// TIA Portal V20 export
// export: Created 2026-10-19T18:41:39.9754622Z, ExportSetting WithDefaults, DisplayName Totally Integrated Automation Portal, DisplayVersion V20 Update 6, DisplayName TIA Portal Openness, DisplayVersion V20 Update 6, DisplayName TIA Portal Version Control Interface, DisplayVersion V20 Update 6, DisplayName SINAMICS Startdrive Advanced, DisplayVersion V20 SP1, DisplayName SINAMICS Startdrive G130, G150, S120, S150, SINAMICS MV, G220, S200, S210, DisplayVersion V20 SP1, DisplayName SINAMICS Startdrive G110M, G120, G120C, G120D, G120P, G115D, DisplayVersion V20 SP1, DisplayName STEP 7 Professional, DisplayVersion V20 Update 6, DisplayName STEP 7 Safety, DisplayVersion V20 Update 2, DisplayName WinCC Basic/Comfort/Advanced, DisplayVersion V20 Update 6, DisplayName WinCC Unified, DisplayVersion V20 Update 6
FUNCTION "FC_CLOCK" : DTL   // FC55, LAD
{ S7_Optimized_Access := 'TRUE' }
VERSION : 0.1
// stored: AutoNumber true, IsIECCheckEnabled false, SetENOAutomatically false, UDAEnableTagReadback false
   VAR_OUTPUT
      CurrentTime : String;
   END_VAR
   VAR_TEMP
      CurrentDTL : DTL;
      RetVal : Int;
      TempString : String;
      strYear : String;
      strMonth : String;
      strDay : String;
      strHour : String;
      strMinute : String;
      strSeconds : String;
   END_VAR
   VAR_TEMP   // added for the SCL form of the ladder/FBD networks
      _w1 : Bool;
      _w2 : Bool;
      _w3 : Bool;
      _w4 : Bool;
      _w5 : Bool;
   END_VAR
BEGIN

REGION Network 1: Read Current Local Time
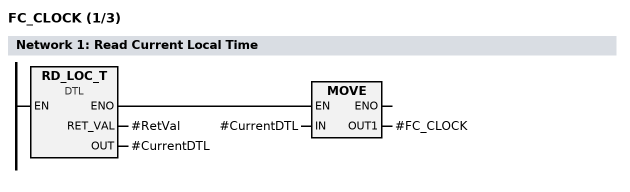
   RUNG wire#powerrail
      { S7_Templates := "date_type := DTL" } RD_LOC_T(RET_VAL => #RetVal, OUT => #CurrentDTL)
      Move(in := #CurrentDTL, out1 => #FC_CLOCK)
   END_RUNG
   // the same network as SCL:
   #RetVal := RD_LOC_T(OUT => #CurrentDTL, ENO => #_w1);
   IF #_w1 THEN #FC_CLOCK := #CurrentDTL; END_IF;
END_REGION

REGION Network 2: Converstion all data to string
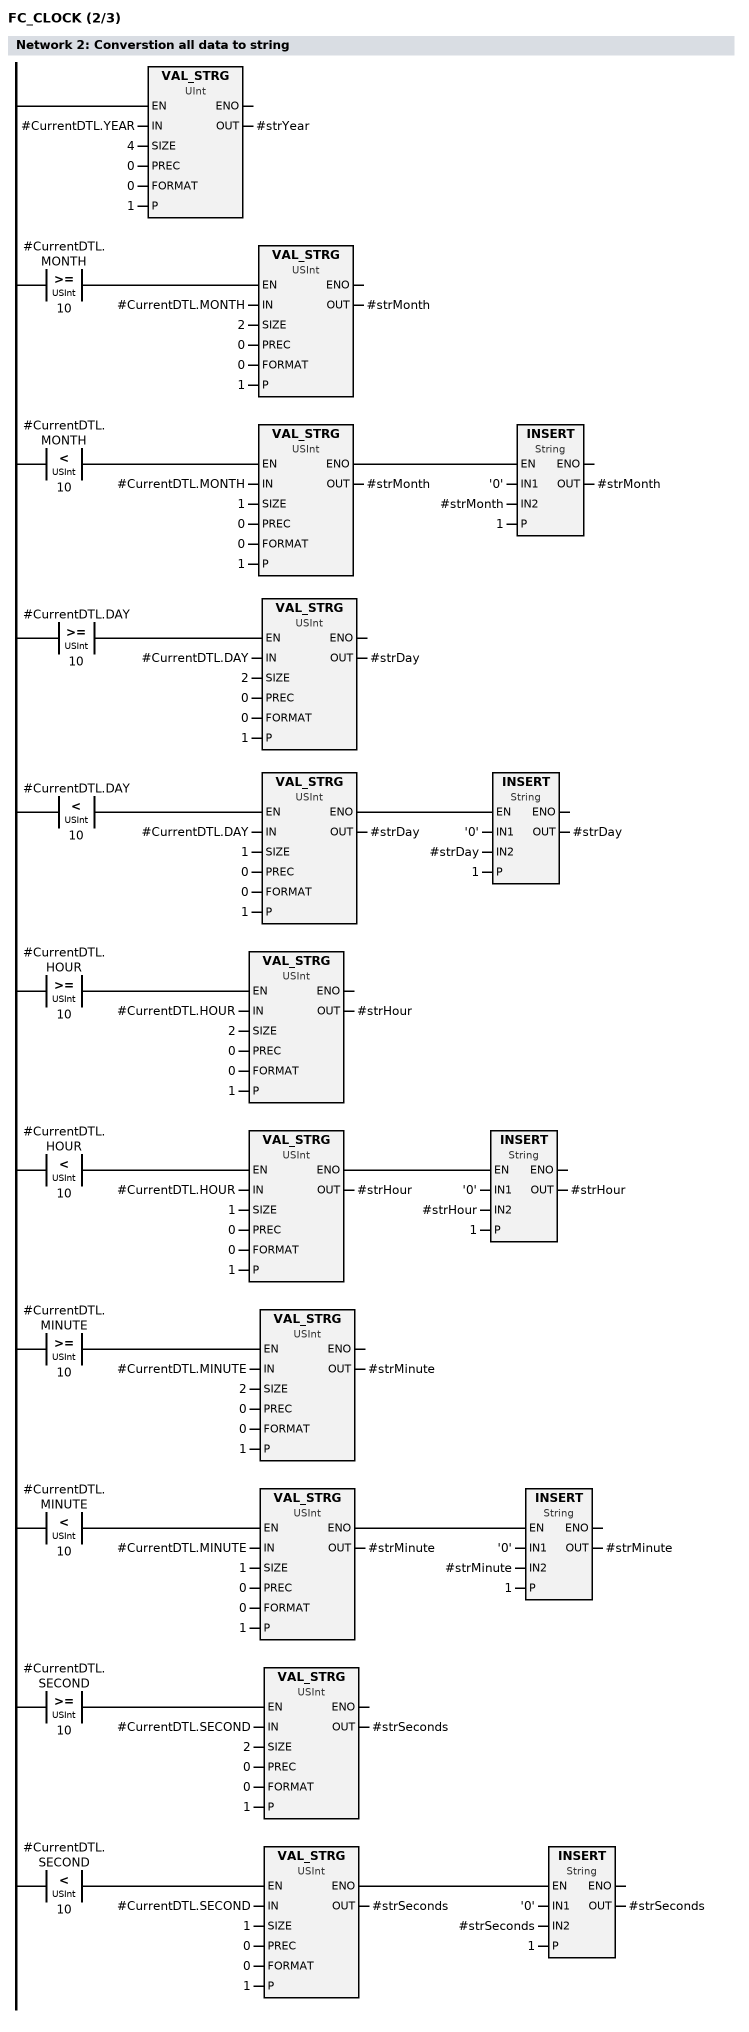
   RUNG wire#powerrail
      { S7_Templates := "[value_type := UInt, str_type := String]" } VAL_STRG(IN := #CurrentDTL.YEAR, SIZE := 4, PREC := 0, FORMAT := 0, P := 1, OUT => #strYear)
   END_RUNG
   RUNG wire#powerrail
      { S7_Templates := "SrcType := USInt" } GE_Contact(in1 := #CurrentDTL.MONTH, in2 := 10)
      { S7_Templates := "[value_type := USInt, str_type := String]" } VAL_STRG(IN := #CurrentDTL.MONTH, SIZE := 2, PREC := 0, FORMAT := 0, P := 1, OUT => #strMonth)
   END_RUNG
   RUNG wire#powerrail
      { S7_Templates := "SrcType := USInt" } LT_Contact(in1 := #CurrentDTL.MONTH, in2 := 10)
      { S7_Templates := "[value_type := USInt, str_type := String]" } VAL_STRG(IN := #CurrentDTL.MONTH, SIZE := 1, PREC := 0, FORMAT := 0, P := 1, OUT => #strMonth)
      { S7_Templates := "str_type := String" } INSERT(IN1 := '0', IN2 := #strMonth, P := 1, OUT => #strMonth)
   END_RUNG
   RUNG wire#powerrail
      { S7_Templates := "SrcType := USInt" } GE_Contact(in1 := #CurrentDTL.DAY, in2 := 10)
      { S7_Templates := "[value_type := USInt, str_type := String]" } VAL_STRG(IN := #CurrentDTL.DAY, SIZE := 2, PREC := 0, FORMAT := 0, P := 1, OUT => #strDay)
   END_RUNG
   RUNG wire#powerrail
      { S7_Templates := "SrcType := USInt" } LT_Contact(in1 := #CurrentDTL.DAY, in2 := 10)
      { S7_Templates := "[value_type := USInt, str_type := String]" } VAL_STRG(IN := #CurrentDTL.DAY, SIZE := 1, PREC := 0, FORMAT := 0, P := 1, OUT => #strDay)
      { S7_Templates := "str_type := String" } INSERT(IN1 := '0', IN2 := #strDay, P := 1, OUT => #strDay)
   END_RUNG
   RUNG wire#powerrail
      { S7_Templates := "SrcType := USInt" } GE_Contact(in1 := #CurrentDTL.HOUR, in2 := 10)
      { S7_Templates := "[value_type := USInt, str_type := String]" } VAL_STRG(IN := #CurrentDTL.HOUR, SIZE := 2, PREC := 0, FORMAT := 0, P := 1, OUT => #strHour)
   END_RUNG
   RUNG wire#powerrail
      { S7_Templates := "SrcType := USInt" } LT_Contact(in1 := #CurrentDTL.HOUR, in2 := 10)
      { S7_Templates := "[value_type := USInt, str_type := String]" } VAL_STRG(IN := #CurrentDTL.HOUR, SIZE := 1, PREC := 0, FORMAT := 0, P := 1, OUT => #strHour)
      { S7_Templates := "str_type := String" } INSERT(IN1 := '0', IN2 := #strHour, P := 1, OUT => #strHour)
   END_RUNG
   RUNG wire#powerrail
      { S7_Templates := "SrcType := USInt" } GE_Contact(in1 := #CurrentDTL.MINUTE, in2 := 10)
      { S7_Templates := "[value_type := USInt, str_type := String]" } VAL_STRG(IN := #CurrentDTL.MINUTE, SIZE := 2, PREC := 0, FORMAT := 0, P := 1, OUT => #strMinute)
   END_RUNG
   RUNG wire#powerrail
      { S7_Templates := "SrcType := USInt" } LT_Contact(in1 := #CurrentDTL.MINUTE, in2 := 10)
      { S7_Templates := "[value_type := USInt, str_type := String]" } VAL_STRG(IN := #CurrentDTL.MINUTE, SIZE := 1, PREC := 0, FORMAT := 0, P := 1, OUT => #strMinute)
      { S7_Templates := "str_type := String" } INSERT(IN1 := '0', IN2 := #strMinute, P := 1, OUT => #strMinute)
   END_RUNG
   RUNG wire#powerrail
      { S7_Templates := "SrcType := USInt" } GE_Contact(in1 := #CurrentDTL.SECOND, in2 := 10)
      { S7_Templates := "[value_type := USInt, str_type := String]" } VAL_STRG(IN := #CurrentDTL.SECOND, SIZE := 2, PREC := 0, FORMAT := 0, P := 1, OUT => #strSeconds)
   END_RUNG
   RUNG wire#powerrail
      { S7_Templates := "SrcType := USInt" } LT_Contact(in1 := #CurrentDTL.SECOND, in2 := 10)
      { S7_Templates := "[value_type := USInt, str_type := String]" } VAL_STRG(IN := #CurrentDTL.SECOND, SIZE := 1, PREC := 0, FORMAT := 0, P := 1, OUT => #strSeconds)
      { S7_Templates := "str_type := String" } INSERT(IN1 := '0', IN2 := #strSeconds, P := 1, OUT => #strSeconds)
   END_RUNG
   // the same network as SCL:
   VAL_STRG(IN := #CurrentDTL.YEAR, SIZE := 4, PREC := 0, FORMAT := 0, P := 1, OUT => #strYear);
   IF #CurrentDTL.MONTH >= 10 THEN
       VAL_STRG(IN := #CurrentDTL.MONTH, SIZE := 2, PREC := 0, FORMAT := 0, P := 1, OUT => #strMonth);
   END_IF;
   VAL_STRG(EN := #CurrentDTL.MONTH < 10,
            IN := #CurrentDTL.MONTH,
            SIZE := 1,
            PREC := 0,
            FORMAT := 0,
            P := 1,
            OUT => #strMonth,
            ENO => #_w1);
   IF #_w1 THEN INSERT(IN1 := '0', IN2 := #strMonth, P := 1, OUT => #strMonth); END_IF;
   IF #CurrentDTL.DAY >= 10 THEN
       VAL_STRG(IN := #CurrentDTL.DAY, SIZE := 2, PREC := 0, FORMAT := 0, P := 1, OUT => #strDay);
   END_IF;
   VAL_STRG(EN := #CurrentDTL.DAY < 10,
            IN := #CurrentDTL.DAY,
            SIZE := 1,
            PREC := 0,
            FORMAT := 0,
            P := 1,
            OUT => #strDay,
            ENO => #_w2);
   IF #_w2 THEN INSERT(IN1 := '0', IN2 := #strDay, P := 1, OUT => #strDay); END_IF;
   IF #CurrentDTL.HOUR >= 10 THEN
       VAL_STRG(IN := #CurrentDTL.HOUR, SIZE := 2, PREC := 0, FORMAT := 0, P := 1, OUT => #strHour);
   END_IF;
   VAL_STRG(EN := #CurrentDTL.HOUR < 10,
            IN := #CurrentDTL.HOUR,
            SIZE := 1,
            PREC := 0,
            FORMAT := 0,
            P := 1,
            OUT => #strHour,
            ENO => #_w3);
   IF #_w3 THEN INSERT(IN1 := '0', IN2 := #strHour, P := 1, OUT => #strHour); END_IF;
   IF #CurrentDTL.MINUTE >= 10 THEN
       VAL_STRG(IN := #CurrentDTL.MINUTE, SIZE := 2, PREC := 0, FORMAT := 0, P := 1, OUT => #strMinute);
   END_IF;
   VAL_STRG(EN := #CurrentDTL.MINUTE < 10,
            IN := #CurrentDTL.MINUTE,
            SIZE := 1,
            PREC := 0,
            FORMAT := 0,
            P := 1,
            OUT => #strMinute,
            ENO => #_w4);
   IF #_w4 THEN INSERT(IN1 := '0', IN2 := #strMinute, P := 1, OUT => #strMinute); END_IF;
   IF #CurrentDTL.SECOND >= 10 THEN
       VAL_STRG(IN := #CurrentDTL.SECOND, SIZE := 2, PREC := 0, FORMAT := 0, P := 1, OUT => #strSeconds);
   END_IF;
   VAL_STRG(EN := #CurrentDTL.SECOND < 10,
            IN := #CurrentDTL.SECOND,
            SIZE := 1,
            PREC := 0,
            FORMAT := 0,
            P := 1,
            OUT => #strSeconds,
            ENO => #_w5);
   IF #_w5 THEN INSERT(IN1 := '0', IN2 := #strSeconds, P := 1, OUT => #strSeconds); END_IF;
END_REGION

REGION Network 3: Current Time String
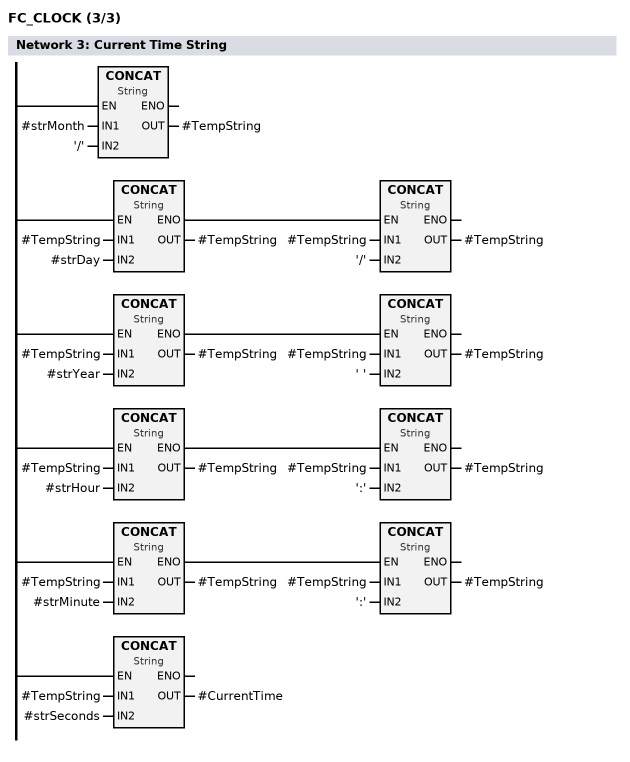
   RUNG wire#powerrail
      { S7_Templates := "[card := 2, str_type := String]" } CONCAT(IN1 := #strMonth, IN2 := '/', OUT => #TempString)
   END_RUNG
   RUNG wire#powerrail
      { S7_Templates := "[card := 2, str_type := String]" } CONCAT(IN1 := #TempString, IN2 := #strDay, OUT => #TempString)
      { S7_Templates := "[card := 2, str_type := String]" } CONCAT(IN1 := #TempString, IN2 := '/', OUT => #TempString)
   END_RUNG
   RUNG wire#powerrail
      { S7_Templates := "[card := 2, str_type := String]" } CONCAT(IN1 := #TempString, IN2 := #strYear, OUT => #TempString)
      { S7_Templates := "[card := 2, str_type := String]" } CONCAT(IN1 := #TempString, IN2 := ' ', OUT => #TempString)
   END_RUNG
   RUNG wire#powerrail
      { S7_Templates := "[card := 2, str_type := String]" } CONCAT(IN1 := #TempString, IN2 := #strHour, OUT => #TempString)
      { S7_Templates := "[card := 2, str_type := String]" } CONCAT(IN1 := #TempString, IN2 := ':', OUT => #TempString)
   END_RUNG
   RUNG wire#powerrail
      { S7_Templates := "[card := 2, str_type := String]" } CONCAT(IN1 := #TempString, IN2 := #strMinute, OUT => #TempString)
      { S7_Templates := "[card := 2, str_type := String]" } CONCAT(IN1 := #TempString, IN2 := ':', OUT => #TempString)
   END_RUNG
   RUNG wire#powerrail
      { S7_Templates := "[card := 2, str_type := String]" } CONCAT(IN1 := #TempString, IN2 := #strSeconds, OUT => #CurrentTime)
   END_RUNG
   // the same network as SCL:
   CONCAT(IN1 := #strMonth, IN2 := '/', OUT => #TempString);
   CONCAT(IN1 := #TempString, IN2 := #strDay, OUT => #TempString, ENO => #_w1);
   IF #_w1 THEN CONCAT(IN1 := #TempString, IN2 := '/', OUT => #TempString); END_IF;
   CONCAT(IN1 := #TempString, IN2 := #strYear, OUT => #TempString, ENO => #_w2);
   IF #_w2 THEN CONCAT(IN1 := #TempString, IN2 := ' ', OUT => #TempString); END_IF;
   CONCAT(IN1 := #TempString, IN2 := #strHour, OUT => #TempString, ENO => #_w3);
   IF #_w3 THEN CONCAT(IN1 := #TempString, IN2 := ':', OUT => #TempString); END_IF;
   CONCAT(IN1 := #TempString, IN2 := #strMinute, OUT => #TempString, ENO => #_w4);
   IF #_w4 THEN CONCAT(IN1 := #TempString, IN2 := ':', OUT => #TempString); END_IF;
   CONCAT(IN1 := #TempString, IN2 := #strSeconds, OUT => #CurrentTime);
END_REGION
END_FUNCTION
